(* IEC 61131-3 sources: STAR-PLC-Agent/results/raw/batch_fresh_20261114/PUB003/functional/attempt_0001, 1 file *)

(* ---- test_program.st ---- *)
PROGRAM PLC_PRG
VAR
 BenchStep : UDINT := 0;
 BenchCalls : UDINT := 0;
 BenchDone : BOOL := FALSE;
 BenchUut0 : FB_Task;
 BenchUut1 : FB_Task;
 BenchUut2 : FB_Task;
 BenchUut3 : FB_Task;
 BenchUut4 : FB_Task;
 BenchUut5 : FB_Task;
 BenchUut6 : FB_Task;
 BenchUut7 : FB_Task;
 TraceIn_Value : ARRAY[0..48] OF REAL;
 TraceIn_hiLevel : ARRAY[0..48] OF REAL;
 TraceIn_loLevel : ARRAY[0..48] OF REAL;
 TraceIn_hystWindow : ARRAY[0..48] OF REAL;
 TraceOut_hiAlarm : ARRAY[0..48] OF BOOL;
 TraceOut_loAlarm : ARRAY[0..48] OF BOOL;
 TraceOut_error : ARRAY[0..48] OF BOOL;
 TraceOut_status : ARRAY[0..48] OF WORD;
END_VAR

IF NOT BenchDone THEN
 CASE BenchStep OF
 0:
   BenchUut0.Value := REAL#50.0;
   BenchUut0.hiLevel := REAL#80.0;
   BenchUut0.loLevel := REAL#20.0;
   BenchUut0.hystWindow := REAL#5.0;
   TraceIn_Value[0] := BenchUut0.Value;
   TraceIn_hiLevel[0] := BenchUut0.hiLevel;
   TraceIn_loLevel[0] := BenchUut0.loLevel;
   TraceIn_hystWindow[0] := BenchUut0.hystWindow;
   BenchUut0();
   TraceOut_hiAlarm[0] := BenchUut0.hiAlarm;
   TraceOut_loAlarm[0] := BenchUut0.loAlarm;
   TraceOut_error[0] := BenchUut0.error;
   TraceOut_status[0] := BenchUut0.status;
   BenchCalls := BenchCalls + 1;
 1:
   BenchUut0.Value := REAL#80.0;
   BenchUut0.hiLevel := REAL#80.0;
   BenchUut0.loLevel := REAL#20.0;
   BenchUut0.hystWindow := REAL#5.0;
   TraceIn_Value[1] := BenchUut0.Value;
   TraceIn_hiLevel[1] := BenchUut0.hiLevel;
   TraceIn_loLevel[1] := BenchUut0.loLevel;
   TraceIn_hystWindow[1] := BenchUut0.hystWindow;
   BenchUut0();
   TraceOut_hiAlarm[1] := BenchUut0.hiAlarm;
   TraceOut_loAlarm[1] := BenchUut0.loAlarm;
   TraceOut_error[1] := BenchUut0.error;
   TraceOut_status[1] := BenchUut0.status;
   BenchCalls := BenchCalls + 1;
 2:
   BenchUut0.Value := REAL#81.0;
   BenchUut0.hiLevel := REAL#80.0;
   BenchUut0.loLevel := REAL#20.0;
   BenchUut0.hystWindow := REAL#5.0;
   TraceIn_Value[2] := BenchUut0.Value;
   TraceIn_hiLevel[2] := BenchUut0.hiLevel;
   TraceIn_loLevel[2] := BenchUut0.loLevel;
   TraceIn_hystWindow[2] := BenchUut0.hystWindow;
   BenchUut0();
   TraceOut_hiAlarm[2] := BenchUut0.hiAlarm;
   TraceOut_loAlarm[2] := BenchUut0.loAlarm;
   TraceOut_error[2] := BenchUut0.error;
   TraceOut_status[2] := BenchUut0.status;
   BenchCalls := BenchCalls + 1;
 3:
   BenchUut0.Value := REAL#75.0;
   BenchUut0.hiLevel := REAL#80.0;
   BenchUut0.loLevel := REAL#20.0;
   BenchUut0.hystWindow := REAL#5.0;
   TraceIn_Value[3] := BenchUut0.Value;
   TraceIn_hiLevel[3] := BenchUut0.hiLevel;
   TraceIn_loLevel[3] := BenchUut0.loLevel;
   TraceIn_hystWindow[3] := BenchUut0.hystWindow;
   BenchUut0();
   TraceOut_hiAlarm[3] := BenchUut0.hiAlarm;
   TraceOut_loAlarm[3] := BenchUut0.loAlarm;
   TraceOut_error[3] := BenchUut0.error;
   TraceOut_status[3] := BenchUut0.status;
   BenchCalls := BenchCalls + 1;
 4:
   BenchUut0.Value := REAL#74.0;
   BenchUut0.hiLevel := REAL#80.0;
   BenchUut0.loLevel := REAL#20.0;
   BenchUut0.hystWindow := REAL#5.0;
   TraceIn_Value[4] := BenchUut0.Value;
   TraceIn_hiLevel[4] := BenchUut0.hiLevel;
   TraceIn_loLevel[4] := BenchUut0.loLevel;
   TraceIn_hystWindow[4] := BenchUut0.hystWindow;
   BenchUut0();
   TraceOut_hiAlarm[4] := BenchUut0.hiAlarm;
   TraceOut_loAlarm[4] := BenchUut0.loAlarm;
   TraceOut_error[4] := BenchUut0.error;
   TraceOut_status[4] := BenchUut0.status;
   BenchCalls := BenchCalls + 1;
 5:
   BenchUut0.Value := REAL#20.0;
   BenchUut0.hiLevel := REAL#80.0;
   BenchUut0.loLevel := REAL#20.0;
   BenchUut0.hystWindow := REAL#5.0;
   TraceIn_Value[5] := BenchUut0.Value;
   TraceIn_hiLevel[5] := BenchUut0.hiLevel;
   TraceIn_loLevel[5] := BenchUut0.loLevel;
   TraceIn_hystWindow[5] := BenchUut0.hystWindow;
   BenchUut0();
   TraceOut_hiAlarm[5] := BenchUut0.hiAlarm;
   TraceOut_loAlarm[5] := BenchUut0.loAlarm;
   TraceOut_error[5] := BenchUut0.error;
   TraceOut_status[5] := BenchUut0.status;
   BenchCalls := BenchCalls + 1;
 6:
   BenchUut0.Value := REAL#19.0;
   BenchUut0.hiLevel := REAL#80.0;
   BenchUut0.loLevel := REAL#20.0;
   BenchUut0.hystWindow := REAL#5.0;
   TraceIn_Value[6] := BenchUut0.Value;
   TraceIn_hiLevel[6] := BenchUut0.hiLevel;
   TraceIn_loLevel[6] := BenchUut0.loLevel;
   TraceIn_hystWindow[6] := BenchUut0.hystWindow;
   BenchUut0();
   TraceOut_hiAlarm[6] := BenchUut0.hiAlarm;
   TraceOut_loAlarm[6] := BenchUut0.loAlarm;
   TraceOut_error[6] := BenchUut0.error;
   TraceOut_status[6] := BenchUut0.status;
   BenchCalls := BenchCalls + 1;
 7:
   BenchUut0.Value := REAL#25.0;
   BenchUut0.hiLevel := REAL#80.0;
   BenchUut0.loLevel := REAL#20.0;
   BenchUut0.hystWindow := REAL#5.0;
   TraceIn_Value[7] := BenchUut0.Value;
   TraceIn_hiLevel[7] := BenchUut0.hiLevel;
   TraceIn_loLevel[7] := BenchUut0.loLevel;
   TraceIn_hystWindow[7] := BenchUut0.hystWindow;
   BenchUut0();
   TraceOut_hiAlarm[7] := BenchUut0.hiAlarm;
   TraceOut_loAlarm[7] := BenchUut0.loAlarm;
   TraceOut_error[7] := BenchUut0.error;
   TraceOut_status[7] := BenchUut0.status;
   BenchCalls := BenchCalls + 1;
 8:
   BenchUut0.Value := REAL#26.0;
   BenchUut0.hiLevel := REAL#80.0;
   BenchUut0.loLevel := REAL#20.0;
   BenchUut0.hystWindow := REAL#5.0;
   TraceIn_Value[8] := BenchUut0.Value;
   TraceIn_hiLevel[8] := BenchUut0.hiLevel;
   TraceIn_loLevel[8] := BenchUut0.loLevel;
   TraceIn_hystWindow[8] := BenchUut0.hystWindow;
   BenchUut0();
   TraceOut_hiAlarm[8] := BenchUut0.hiAlarm;
   TraceOut_loAlarm[8] := BenchUut0.loAlarm;
   TraceOut_error[8] := BenchUut0.error;
   TraceOut_status[8] := BenchUut0.status;
   BenchCalls := BenchCalls + 1;
 9:
   BenchUut1.Value := REAL#90.0;
   BenchUut1.hiLevel := REAL#80.0;
   BenchUut1.loLevel := REAL#20.0;
   BenchUut1.hystWindow := REAL#5.0;
   TraceIn_Value[9] := BenchUut1.Value;
   TraceIn_hiLevel[9] := BenchUut1.hiLevel;
   TraceIn_loLevel[9] := BenchUut1.loLevel;
   TraceIn_hystWindow[9] := BenchUut1.hystWindow;
   BenchUut1();
   TraceOut_hiAlarm[9] := BenchUut1.hiAlarm;
   TraceOut_loAlarm[9] := BenchUut1.loAlarm;
   TraceOut_error[9] := BenchUut1.error;
   TraceOut_status[9] := BenchUut1.status;
   BenchCalls := BenchCalls + 1;
 10:
   BenchUut1.Value := REAL#50.0;
   BenchUut1.hiLevel := REAL#80.0;
   BenchUut1.loLevel := REAL#80.0;
   BenchUut1.hystWindow := REAL#80.0;
   TraceIn_Value[10] := BenchUut1.Value;
   TraceIn_hiLevel[10] := BenchUut1.hiLevel;
   TraceIn_loLevel[10] := BenchUut1.loLevel;
   TraceIn_hystWindow[10] := BenchUut1.hystWindow;
   BenchUut1();
   TraceOut_hiAlarm[10] := BenchUut1.hiAlarm;
   TraceOut_loAlarm[10] := BenchUut1.loAlarm;
   TraceOut_error[10] := BenchUut1.error;
   TraceOut_status[10] := BenchUut1.status;
   BenchCalls := BenchCalls + 1;
 11:
   BenchUut1.Value := REAL#50.0;
   BenchUut1.hiLevel := REAL#80.0;
   BenchUut1.loLevel := REAL#20.0;
   BenchUut1.hystWindow := REAL#60.0;
   TraceIn_Value[11] := BenchUut1.Value;
   TraceIn_hiLevel[11] := BenchUut1.hiLevel;
   TraceIn_loLevel[11] := BenchUut1.loLevel;
   TraceIn_hystWindow[11] := BenchUut1.hystWindow;
   BenchUut1();
   TraceOut_hiAlarm[11] := BenchUut1.hiAlarm;
   TraceOut_loAlarm[11] := BenchUut1.loAlarm;
   TraceOut_error[11] := BenchUut1.error;
   TraceOut_status[11] := BenchUut1.status;
   BenchCalls := BenchCalls + 1;
 12:
   BenchUut1.Value := REAL#50.0;
   BenchUut1.hiLevel := REAL#80.0;
   BenchUut1.loLevel := REAL#20.0;
   BenchUut1.hystWindow := REAL#5.0;
   TraceIn_Value[12] := BenchUut1.Value;
   TraceIn_hiLevel[12] := BenchUut1.hiLevel;
   TraceIn_loLevel[12] := BenchUut1.loLevel;
   TraceIn_hystWindow[12] := BenchUut1.hystWindow;
   BenchUut1();
   TraceOut_hiAlarm[12] := BenchUut1.hiAlarm;
   TraceOut_loAlarm[12] := BenchUut1.loAlarm;
   TraceOut_error[12] := BenchUut1.error;
   TraceOut_status[12] := BenchUut1.status;
   BenchCalls := BenchCalls + 1;
 13:
   BenchUut2.Value := REAL#101.0;
   BenchUut2.hiLevel := REAL#100.0;
   BenchUut2.loLevel := REAL#0.0;
   BenchUut2.hystWindow := REAL#90.0;
   TraceIn_Value[13] := BenchUut2.Value;
   TraceIn_hiLevel[13] := BenchUut2.hiLevel;
   TraceIn_loLevel[13] := BenchUut2.loLevel;
   TraceIn_hystWindow[13] := BenchUut2.hystWindow;
   BenchUut2();
   TraceOut_hiAlarm[13] := BenchUut2.hiAlarm;
   TraceOut_loAlarm[13] := BenchUut2.loAlarm;
   TraceOut_error[13] := BenchUut2.error;
   TraceOut_status[13] := BenchUut2.status;
   BenchCalls := BenchCalls + 1;
 14:
   BenchUut2.Value := REAL#50.0;
   BenchUut2.hiLevel := REAL#100.0;
   BenchUut2.loLevel := REAL#0.0;
   BenchUut2.hystWindow := REAL#90.0;
   TraceIn_Value[14] := BenchUut2.Value;
   TraceIn_hiLevel[14] := BenchUut2.hiLevel;
   TraceIn_loLevel[14] := BenchUut2.loLevel;
   TraceIn_hystWindow[14] := BenchUut2.hystWindow;
   BenchUut2();
   TraceOut_hiAlarm[14] := BenchUut2.hiAlarm;
   TraceOut_loAlarm[14] := BenchUut2.loAlarm;
   TraceOut_error[14] := BenchUut2.error;
   TraceOut_status[14] := BenchUut2.status;
   BenchCalls := BenchCalls + 1;
 15:
   BenchUut2.Value := REAL#50.0;
   BenchUut2.hiLevel := REAL#100.0;
   BenchUut2.loLevel := REAL#100.0;
   BenchUut2.hystWindow := REAL#90.0;
   TraceIn_Value[15] := BenchUut2.Value;
   TraceIn_hiLevel[15] := BenchUut2.hiLevel;
   TraceIn_loLevel[15] := BenchUut2.loLevel;
   TraceIn_hystWindow[15] := BenchUut2.hystWindow;
   BenchUut2();
   TraceOut_hiAlarm[15] := BenchUut2.hiAlarm;
   TraceOut_loAlarm[15] := BenchUut2.loAlarm;
   TraceOut_error[15] := BenchUut2.error;
   TraceOut_status[15] := BenchUut2.status;
   BenchCalls := BenchCalls + 1;
 16:
   BenchUut2.Value := REAL#10.0;
   BenchUut2.hiLevel := REAL#100.0;
   BenchUut2.loLevel := REAL#0.0;
   BenchUut2.hystWindow := REAL#90.0;
   TraceIn_Value[16] := BenchUut2.Value;
   TraceIn_hiLevel[16] := BenchUut2.hiLevel;
   TraceIn_loLevel[16] := BenchUut2.loLevel;
   TraceIn_hystWindow[16] := BenchUut2.hystWindow;
   BenchUut2();
   TraceOut_hiAlarm[16] := BenchUut2.hiAlarm;
   TraceOut_loAlarm[16] := BenchUut2.loAlarm;
   TraceOut_error[16] := BenchUut2.error;
   TraceOut_status[16] := BenchUut2.status;
   BenchCalls := BenchCalls + 1;
 17:
   BenchUut2.Value := REAL#9.0;
   BenchUut2.hiLevel := REAL#100.0;
   BenchUut2.loLevel := REAL#0.0;
   BenchUut2.hystWindow := REAL#90.0;
   TraceIn_Value[17] := BenchUut2.Value;
   TraceIn_hiLevel[17] := BenchUut2.hiLevel;
   TraceIn_loLevel[17] := BenchUut2.loLevel;
   TraceIn_hystWindow[17] := BenchUut2.hystWindow;
   BenchUut2();
   TraceOut_hiAlarm[17] := BenchUut2.hiAlarm;
   TraceOut_loAlarm[17] := BenchUut2.loAlarm;
   TraceOut_error[17] := BenchUut2.error;
   TraceOut_status[17] := BenchUut2.status;
   BenchCalls := BenchCalls + 1;
 18:
   BenchUut2.Value := REAL#-1.0;
   BenchUut2.hiLevel := REAL#100.0;
   BenchUut2.loLevel := REAL#0.0;
   BenchUut2.hystWindow := REAL#90.0;
   TraceIn_Value[18] := BenchUut2.Value;
   TraceIn_hiLevel[18] := BenchUut2.hiLevel;
   TraceIn_loLevel[18] := BenchUut2.loLevel;
   TraceIn_hystWindow[18] := BenchUut2.hystWindow;
   BenchUut2();
   TraceOut_hiAlarm[18] := BenchUut2.hiAlarm;
   TraceOut_loAlarm[18] := BenchUut2.loAlarm;
   TraceOut_error[18] := BenchUut2.error;
   TraceOut_status[18] := BenchUut2.status;
   BenchCalls := BenchCalls + 1;
 19:
   BenchUut3.Value := REAL#5.0;
   BenchUut3.hiLevel := REAL#50.0;
   BenchUut3.loLevel := REAL#10.0;
   BenchUut3.hystWindow := REAL#5.0;
   TraceIn_Value[19] := BenchUut3.Value;
   TraceIn_hiLevel[19] := BenchUut3.hiLevel;
   TraceIn_loLevel[19] := BenchUut3.loLevel;
   TraceIn_hystWindow[19] := BenchUut3.hystWindow;
   BenchUut3();
   TraceOut_hiAlarm[19] := BenchUut3.hiAlarm;
   TraceOut_loAlarm[19] := BenchUut3.loAlarm;
   TraceOut_error[19] := BenchUut3.error;
   TraceOut_status[19] := BenchUut3.status;
   BenchCalls := BenchCalls + 1;
 20:
   BenchUut3.Value := REAL#25.0;
   BenchUut3.hiLevel := REAL#50.0;
   BenchUut3.loLevel := REAL#60.0;
   BenchUut3.hystWindow := REAL#5.0;
   TraceIn_Value[20] := BenchUut3.Value;
   TraceIn_hiLevel[20] := BenchUut3.hiLevel;
   TraceIn_loLevel[20] := BenchUut3.loLevel;
   TraceIn_hystWindow[20] := BenchUut3.hystWindow;
   BenchUut3();
   TraceOut_hiAlarm[20] := BenchUut3.hiAlarm;
   TraceOut_loAlarm[20] := BenchUut3.loAlarm;
   TraceOut_error[20] := BenchUut3.error;
   TraceOut_status[20] := BenchUut3.status;
   BenchCalls := BenchCalls + 1;
 21:
   BenchUut3.Value := REAL#25.0;
   BenchUut3.hiLevel := REAL#50.0;
   BenchUut3.loLevel := REAL#10.0;
   BenchUut3.hystWindow := REAL#40.0;
   TraceIn_Value[21] := BenchUut3.Value;
   TraceIn_hiLevel[21] := BenchUut3.hiLevel;
   TraceIn_loLevel[21] := BenchUut3.loLevel;
   TraceIn_hystWindow[21] := BenchUut3.hystWindow;
   BenchUut3();
   TraceOut_hiAlarm[21] := BenchUut3.hiAlarm;
   TraceOut_loAlarm[21] := BenchUut3.loAlarm;
   TraceOut_error[21] := BenchUut3.error;
   TraceOut_status[21] := BenchUut3.status;
   BenchCalls := BenchCalls + 1;
 22:
   BenchUut3.Value := REAL#16.0;
   BenchUut3.hiLevel := REAL#50.0;
   BenchUut3.loLevel := REAL#10.0;
   BenchUut3.hystWindow := REAL#5.0;
   TraceIn_Value[22] := BenchUut3.Value;
   TraceIn_hiLevel[22] := BenchUut3.hiLevel;
   TraceIn_loLevel[22] := BenchUut3.loLevel;
   TraceIn_hystWindow[22] := BenchUut3.hystWindow;
   BenchUut3();
   TraceOut_hiAlarm[22] := BenchUut3.hiAlarm;
   TraceOut_loAlarm[22] := BenchUut3.loAlarm;
   TraceOut_error[22] := BenchUut3.error;
   TraceOut_status[22] := BenchUut3.status;
   BenchCalls := BenchCalls + 1;
 23:
   BenchUut3.Value := REAL#10.125;
   BenchUut3.hiLevel := REAL#20.375;
   BenchUut3.loLevel := REAL#10.125;
   BenchUut3.hystWindow := REAL#0.0;
   TraceIn_Value[23] := BenchUut3.Value;
   TraceIn_hiLevel[23] := BenchUut3.hiLevel;
   TraceIn_loLevel[23] := BenchUut3.loLevel;
   TraceIn_hystWindow[23] := BenchUut3.hystWindow;
   BenchUut3();
   TraceOut_hiAlarm[23] := BenchUut3.hiAlarm;
   TraceOut_loAlarm[23] := BenchUut3.loAlarm;
   TraceOut_error[23] := BenchUut3.error;
   TraceOut_status[23] := BenchUut3.status;
   BenchCalls := BenchCalls + 1;
 24:
   BenchUut3.Value := REAL#20.3751;
   BenchUut3.hiLevel := REAL#20.375;
   BenchUut3.loLevel := REAL#10.125;
   BenchUut3.hystWindow := REAL#0.0;
   TraceIn_Value[24] := BenchUut3.Value;
   TraceIn_hiLevel[24] := BenchUut3.hiLevel;
   TraceIn_loLevel[24] := BenchUut3.loLevel;
   TraceIn_hystWindow[24] := BenchUut3.hystWindow;
   BenchUut3();
   TraceOut_hiAlarm[24] := BenchUut3.hiAlarm;
   TraceOut_loAlarm[24] := BenchUut3.loAlarm;
   TraceOut_error[24] := BenchUut3.error;
   TraceOut_status[24] := BenchUut3.status;
   BenchCalls := BenchCalls + 1;
 25:
   BenchUut3.Value := REAL#20.25;
   BenchUut3.hiLevel := REAL#20.375;
   BenchUut3.loLevel := REAL#10.125;
   BenchUut3.hystWindow := REAL#0.0;
   TraceIn_Value[25] := BenchUut3.Value;
   TraceIn_hiLevel[25] := BenchUut3.hiLevel;
   TraceIn_loLevel[25] := BenchUut3.loLevel;
   TraceIn_hystWindow[25] := BenchUut3.hystWindow;
   BenchUut3();
   TraceOut_hiAlarm[25] := BenchUut3.hiAlarm;
   TraceOut_loAlarm[25] := BenchUut3.loAlarm;
   TraceOut_error[25] := BenchUut3.error;
   TraceOut_status[25] := BenchUut3.status;
   BenchCalls := BenchCalls + 1;
 26:
   BenchUut4.Value := REAL#19.0;
   BenchUut4.hiLevel := REAL#80.0;
   BenchUut4.loLevel := REAL#20.0;
   BenchUut4.hystWindow := REAL#5.0;
   TraceIn_Value[26] := BenchUut4.Value;
   TraceIn_hiLevel[26] := BenchUut4.hiLevel;
   TraceIn_loLevel[26] := BenchUut4.loLevel;
   TraceIn_hystWindow[26] := BenchUut4.hystWindow;
   BenchUut4();
   TraceOut_hiAlarm[26] := BenchUut4.hiAlarm;
   TraceOut_loAlarm[26] := BenchUut4.loAlarm;
   TraceOut_error[26] := BenchUut4.error;
   TraceOut_status[26] := BenchUut4.status;
   BenchCalls := BenchCalls + 1;
 27:
   BenchUut4.Value := REAL#50.0;
   BenchUut4.hiLevel := REAL#80.0;
   BenchUut4.loLevel := REAL#80.0;
   BenchUut4.hystWindow := REAL#80.0;
   TraceIn_Value[27] := BenchUut4.Value;
   TraceIn_hiLevel[27] := BenchUut4.hiLevel;
   TraceIn_loLevel[27] := BenchUut4.loLevel;
   TraceIn_hystWindow[27] := BenchUut4.hystWindow;
   BenchUut4();
   TraceOut_hiAlarm[27] := BenchUut4.hiAlarm;
   TraceOut_loAlarm[27] := BenchUut4.loAlarm;
   TraceOut_error[27] := BenchUut4.error;
   TraceOut_status[27] := BenchUut4.status;
   BenchCalls := BenchCalls + 1;
 28:
   BenchUut5.Value := REAL#1.1;
   BenchUut5.hiLevel := REAL#1.0;
   BenchUut5.loLevel := REAL#0.0;
   BenchUut5.hystWindow := REAL#0.10000000149011612;
   TraceIn_Value[28] := BenchUut5.Value;
   TraceIn_hiLevel[28] := BenchUut5.hiLevel;
   TraceIn_loLevel[28] := BenchUut5.loLevel;
   TraceIn_hystWindow[28] := BenchUut5.hystWindow;
   BenchUut5();
   TraceOut_hiAlarm[28] := BenchUut5.hiAlarm;
   TraceOut_loAlarm[28] := BenchUut5.loAlarm;
   TraceOut_error[28] := BenchUut5.error;
   TraceOut_status[28] := BenchUut5.status;
   BenchCalls := BenchCalls + 1;
 29:
   BenchUut5.Value := REAL#1.0;
   BenchUut5.hiLevel := REAL#1.0;
   BenchUut5.loLevel := REAL#0.0;
   BenchUut5.hystWindow := REAL#0.10000000149011612;
   TraceIn_Value[29] := BenchUut5.Value;
   TraceIn_hiLevel[29] := BenchUut5.hiLevel;
   TraceIn_loLevel[29] := BenchUut5.loLevel;
   TraceIn_hystWindow[29] := BenchUut5.hystWindow;
   BenchUut5();
   TraceOut_hiAlarm[29] := BenchUut5.hiAlarm;
   TraceOut_loAlarm[29] := BenchUut5.loAlarm;
   TraceOut_error[29] := BenchUut5.error;
   TraceOut_status[29] := BenchUut5.status;
   BenchCalls := BenchCalls + 1;
 30:
   BenchUut5.Value := REAL#0.8999999761581421;
   BenchUut5.hiLevel := REAL#1.0;
   BenchUut5.loLevel := REAL#0.0;
   BenchUut5.hystWindow := REAL#0.10000000149011612;
   TraceIn_Value[30] := BenchUut5.Value;
   TraceIn_hiLevel[30] := BenchUut5.hiLevel;
   TraceIn_loLevel[30] := BenchUut5.loLevel;
   TraceIn_hystWindow[30] := BenchUut5.hystWindow;
   BenchUut5();
   TraceOut_hiAlarm[30] := BenchUut5.hiAlarm;
   TraceOut_loAlarm[30] := BenchUut5.loAlarm;
   TraceOut_error[30] := BenchUut5.error;
   TraceOut_status[30] := BenchUut5.status;
   BenchCalls := BenchCalls + 1;
 31:
   BenchUut5.Value := REAL#0.8999989628791809;
   BenchUut5.hiLevel := REAL#1.0;
   BenchUut5.loLevel := REAL#0.0;
   BenchUut5.hystWindow := REAL#0.10000000149011612;
   TraceIn_Value[31] := BenchUut5.Value;
   TraceIn_hiLevel[31] := BenchUut5.hiLevel;
   TraceIn_loLevel[31] := BenchUut5.loLevel;
   TraceIn_hystWindow[31] := BenchUut5.hystWindow;
   BenchUut5();
   TraceOut_hiAlarm[31] := BenchUut5.hiAlarm;
   TraceOut_loAlarm[31] := BenchUut5.loAlarm;
   TraceOut_error[31] := BenchUut5.error;
   TraceOut_status[31] := BenchUut5.status;
   BenchCalls := BenchCalls + 1;
 32:
   BenchUut5.Value := REAL#-0.1;
   BenchUut5.hiLevel := REAL#1.0;
   BenchUut5.loLevel := REAL#0.0;
   BenchUut5.hystWindow := REAL#0.10000000149011612;
   TraceIn_Value[32] := BenchUut5.Value;
   TraceIn_hiLevel[32] := BenchUut5.hiLevel;
   TraceIn_loLevel[32] := BenchUut5.loLevel;
   TraceIn_hystWindow[32] := BenchUut5.hystWindow;
   BenchUut5();
   TraceOut_hiAlarm[32] := BenchUut5.hiAlarm;
   TraceOut_loAlarm[32] := BenchUut5.loAlarm;
   TraceOut_error[32] := BenchUut5.error;
   TraceOut_status[32] := BenchUut5.status;
   BenchCalls := BenchCalls + 1;
 33:
   BenchUut5.Value := REAL#0.0;
   BenchUut5.hiLevel := REAL#1.0;
   BenchUut5.loLevel := REAL#0.0;
   BenchUut5.hystWindow := REAL#0.10000000149011612;
   TraceIn_Value[33] := BenchUut5.Value;
   TraceIn_hiLevel[33] := BenchUut5.hiLevel;
   TraceIn_loLevel[33] := BenchUut5.loLevel;
   TraceIn_hystWindow[33] := BenchUut5.hystWindow;
   BenchUut5();
   TraceOut_hiAlarm[33] := BenchUut5.hiAlarm;
   TraceOut_loAlarm[33] := BenchUut5.loAlarm;
   TraceOut_error[33] := BenchUut5.error;
   TraceOut_status[33] := BenchUut5.status;
   BenchCalls := BenchCalls + 1;
 34:
   BenchUut5.Value := REAL#0.10000000149011612;
   BenchUut5.hiLevel := REAL#1.0;
   BenchUut5.loLevel := REAL#0.0;
   BenchUut5.hystWindow := REAL#0.10000000149011612;
   TraceIn_Value[34] := BenchUut5.Value;
   TraceIn_hiLevel[34] := BenchUut5.hiLevel;
   TraceIn_loLevel[34] := BenchUut5.loLevel;
   TraceIn_hystWindow[34] := BenchUut5.hystWindow;
   BenchUut5();
   TraceOut_hiAlarm[34] := BenchUut5.hiAlarm;
   TraceOut_loAlarm[34] := BenchUut5.loAlarm;
   TraceOut_error[34] := BenchUut5.error;
   TraceOut_status[34] := BenchUut5.status;
   BenchCalls := BenchCalls + 1;
 35:
   BenchUut5.Value := REAL#0.10000099986791611;
   BenchUut5.hiLevel := REAL#1.0;
   BenchUut5.loLevel := REAL#0.0;
   BenchUut5.hystWindow := REAL#0.10000000149011612;
   TraceIn_Value[35] := BenchUut5.Value;
   TraceIn_hiLevel[35] := BenchUut5.hiLevel;
   TraceIn_loLevel[35] := BenchUut5.loLevel;
   TraceIn_hystWindow[35] := BenchUut5.hystWindow;
   BenchUut5();
   TraceOut_hiAlarm[35] := BenchUut5.hiAlarm;
   TraceOut_loAlarm[35] := BenchUut5.loAlarm;
   TraceOut_error[35] := BenchUut5.error;
   TraceOut_status[35] := BenchUut5.status;
   BenchCalls := BenchCalls + 1;
 36:
   BenchUut6.Value := REAL#-9.0;
   BenchUut6.hiLevel := REAL#-10.0;
   BenchUut6.loLevel := REAL#-50.0;
   BenchUut6.hystWindow := REAL#5.0;
   TraceIn_Value[36] := BenchUut6.Value;
   TraceIn_hiLevel[36] := BenchUut6.hiLevel;
   TraceIn_loLevel[36] := BenchUut6.loLevel;
   TraceIn_hystWindow[36] := BenchUut6.hystWindow;
   BenchUut6();
   TraceOut_hiAlarm[36] := BenchUut6.hiAlarm;
   TraceOut_loAlarm[36] := BenchUut6.loAlarm;
   TraceOut_error[36] := BenchUut6.error;
   TraceOut_status[36] := BenchUut6.status;
   BenchCalls := BenchCalls + 1;
 37:
   BenchUut6.Value := REAL#-15.0;
   BenchUut6.hiLevel := REAL#-10.0;
   BenchUut6.loLevel := REAL#-50.0;
   BenchUut6.hystWindow := REAL#5.0;
   TraceIn_Value[37] := BenchUut6.Value;
   TraceIn_hiLevel[37] := BenchUut6.hiLevel;
   TraceIn_loLevel[37] := BenchUut6.loLevel;
   TraceIn_hystWindow[37] := BenchUut6.hystWindow;
   BenchUut6();
   TraceOut_hiAlarm[37] := BenchUut6.hiAlarm;
   TraceOut_loAlarm[37] := BenchUut6.loAlarm;
   TraceOut_error[37] := BenchUut6.error;
   TraceOut_status[37] := BenchUut6.status;
   BenchCalls := BenchCalls + 1;
 38:
   BenchUut6.Value := REAL#-15.1;
   BenchUut6.hiLevel := REAL#-10.0;
   BenchUut6.loLevel := REAL#-50.0;
   BenchUut6.hystWindow := REAL#5.0;
   TraceIn_Value[38] := BenchUut6.Value;
   TraceIn_hiLevel[38] := BenchUut6.hiLevel;
   TraceIn_loLevel[38] := BenchUut6.loLevel;
   TraceIn_hystWindow[38] := BenchUut6.hystWindow;
   BenchUut6();
   TraceOut_hiAlarm[38] := BenchUut6.hiAlarm;
   TraceOut_loAlarm[38] := BenchUut6.loAlarm;
   TraceOut_error[38] := BenchUut6.error;
   TraceOut_status[38] := BenchUut6.status;
   BenchCalls := BenchCalls + 1;
 39:
   BenchUut6.Value := REAL#-51.0;
   BenchUut6.hiLevel := REAL#-10.0;
   BenchUut6.loLevel := REAL#-50.0;
   BenchUut6.hystWindow := REAL#5.0;
   TraceIn_Value[39] := BenchUut6.Value;
   TraceIn_hiLevel[39] := BenchUut6.hiLevel;
   TraceIn_loLevel[39] := BenchUut6.loLevel;
   TraceIn_hystWindow[39] := BenchUut6.hystWindow;
   BenchUut6();
   TraceOut_hiAlarm[39] := BenchUut6.hiAlarm;
   TraceOut_loAlarm[39] := BenchUut6.loAlarm;
   TraceOut_error[39] := BenchUut6.error;
   TraceOut_status[39] := BenchUut6.status;
   BenchCalls := BenchCalls + 1;
 40:
   BenchUut6.Value := REAL#-45.0;
   BenchUut6.hiLevel := REAL#-10.0;
   BenchUut6.loLevel := REAL#-50.0;
   BenchUut6.hystWindow := REAL#5.0;
   TraceIn_Value[40] := BenchUut6.Value;
   TraceIn_hiLevel[40] := BenchUut6.hiLevel;
   TraceIn_loLevel[40] := BenchUut6.loLevel;
   TraceIn_hystWindow[40] := BenchUut6.hystWindow;
   BenchUut6();
   TraceOut_hiAlarm[40] := BenchUut6.hiAlarm;
   TraceOut_loAlarm[40] := BenchUut6.loAlarm;
   TraceOut_error[40] := BenchUut6.error;
   TraceOut_status[40] := BenchUut6.status;
   BenchCalls := BenchCalls + 1;
 41:
   BenchUut6.Value := REAL#-44.9;
   BenchUut6.hiLevel := REAL#-10.0;
   BenchUut6.loLevel := REAL#-50.0;
   BenchUut6.hystWindow := REAL#5.0;
   TraceIn_Value[41] := BenchUut6.Value;
   TraceIn_hiLevel[41] := BenchUut6.hiLevel;
   TraceIn_loLevel[41] := BenchUut6.loLevel;
   TraceIn_hystWindow[41] := BenchUut6.hystWindow;
   BenchUut6();
   TraceOut_hiAlarm[41] := BenchUut6.hiAlarm;
   TraceOut_loAlarm[41] := BenchUut6.loAlarm;
   TraceOut_error[41] := BenchUut6.error;
   TraceOut_status[41] := BenchUut6.status;
   BenchCalls := BenchCalls + 1;
 42:
   BenchUut6.Value := REAL#0.0;
   BenchUut6.hiLevel := REAL#-10.0;
   BenchUut6.loLevel := REAL#-50.0;
   BenchUut6.hystWindow := REAL#5.0;
   TraceIn_Value[42] := BenchUut6.Value;
   TraceIn_hiLevel[42] := BenchUut6.hiLevel;
   TraceIn_loLevel[42] := BenchUut6.loLevel;
   TraceIn_hystWindow[42] := BenchUut6.hystWindow;
   BenchUut6();
   TraceOut_hiAlarm[42] := BenchUut6.hiAlarm;
   TraceOut_loAlarm[42] := BenchUut6.loAlarm;
   TraceOut_error[42] := BenchUut6.error;
   TraceOut_status[42] := BenchUut6.status;
   BenchCalls := BenchCalls + 1;
 43:
   BenchUut6.Value := REAL#-60.0;
   BenchUut6.hiLevel := REAL#-10.0;
   BenchUut6.loLevel := REAL#-50.0;
   BenchUut6.hystWindow := REAL#5.0;
   TraceIn_Value[43] := BenchUut6.Value;
   TraceIn_hiLevel[43] := BenchUut6.hiLevel;
   TraceIn_loLevel[43] := BenchUut6.loLevel;
   TraceIn_hystWindow[43] := BenchUut6.hystWindow;
   BenchUut6();
   TraceOut_hiAlarm[43] := BenchUut6.hiAlarm;
   TraceOut_loAlarm[43] := BenchUut6.loAlarm;
   TraceOut_error[43] := BenchUut6.error;
   TraceOut_status[43] := BenchUut6.status;
   BenchCalls := BenchCalls + 1;
 44:
   BenchUut7.Value := REAL#85.0;
   BenchUut7.hiLevel := REAL#80.0;
   BenchUut7.loLevel := REAL#20.0;
   BenchUut7.hystWindow := REAL#5.0;
   TraceIn_Value[44] := BenchUut7.Value;
   TraceIn_hiLevel[44] := BenchUut7.hiLevel;
   TraceIn_loLevel[44] := BenchUut7.loLevel;
   TraceIn_hystWindow[44] := BenchUut7.hystWindow;
   BenchUut7();
   TraceOut_hiAlarm[44] := BenchUut7.hiAlarm;
   TraceOut_loAlarm[44] := BenchUut7.loAlarm;
   TraceOut_error[44] := BenchUut7.error;
   TraceOut_status[44] := BenchUut7.status;
   BenchCalls := BenchCalls + 1;
 45:
   BenchUut7.Value := REAL#10.0;
   BenchUut7.hiLevel := REAL#80.0;
   BenchUut7.loLevel := REAL#20.0;
   BenchUut7.hystWindow := REAL#60.0;
   TraceIn_Value[45] := BenchUut7.Value;
   TraceIn_hiLevel[45] := BenchUut7.hiLevel;
   TraceIn_loLevel[45] := BenchUut7.loLevel;
   TraceIn_hystWindow[45] := BenchUut7.hystWindow;
   BenchUut7();
   TraceOut_hiAlarm[45] := BenchUut7.hiAlarm;
   TraceOut_loAlarm[45] := BenchUut7.loAlarm;
   TraceOut_error[45] := BenchUut7.error;
   TraceOut_status[45] := BenchUut7.status;
   BenchCalls := BenchCalls + 1;
 46:
   BenchUut7.Value := REAL#10.0;
   BenchUut7.hiLevel := REAL#50.0;
   BenchUut7.loLevel := REAL#60.0;
   BenchUut7.hystWindow := REAL#5.0;
   TraceIn_Value[46] := BenchUut7.Value;
   TraceIn_hiLevel[46] := BenchUut7.hiLevel;
   TraceIn_loLevel[46] := BenchUut7.loLevel;
   TraceIn_hystWindow[46] := BenchUut7.hystWindow;
   BenchUut7();
   TraceOut_hiAlarm[46] := BenchUut7.hiAlarm;
   TraceOut_loAlarm[46] := BenchUut7.loAlarm;
   TraceOut_error[46] := BenchUut7.error;
   TraceOut_status[46] := BenchUut7.status;
   BenchCalls := BenchCalls + 1;
 47:
   BenchUut7.Value := REAL#75.0;
   BenchUut7.hiLevel := REAL#80.0;
   BenchUut7.loLevel := REAL#20.0;
   BenchUut7.hystWindow := REAL#5.0;
   TraceIn_Value[47] := BenchUut7.Value;
   TraceIn_hiLevel[47] := BenchUut7.hiLevel;
   TraceIn_loLevel[47] := BenchUut7.loLevel;
   TraceIn_hystWindow[47] := BenchUut7.hystWindow;
   BenchUut7();
   TraceOut_hiAlarm[47] := BenchUut7.hiAlarm;
   TraceOut_loAlarm[47] := BenchUut7.loAlarm;
   TraceOut_error[47] := BenchUut7.error;
   TraceOut_status[47] := BenchUut7.status;
   BenchCalls := BenchCalls + 1;
 48:
   BenchUut7.Value := REAL#74.0;
   BenchUut7.hiLevel := REAL#80.0;
   BenchUut7.loLevel := REAL#20.0;
   BenchUut7.hystWindow := REAL#5.0;
   TraceIn_Value[48] := BenchUut7.Value;
   TraceIn_hiLevel[48] := BenchUut7.hiLevel;
   TraceIn_loLevel[48] := BenchUut7.loLevel;
   TraceIn_hystWindow[48] := BenchUut7.hystWindow;
   BenchUut7();
   TraceOut_hiAlarm[48] := BenchUut7.hiAlarm;
   TraceOut_loAlarm[48] := BenchUut7.loAlarm;
   TraceOut_error[48] := BenchUut7.error;
   TraceOut_status[48] := BenchUut7.status;
   BenchCalls := BenchCalls + 1;
 END_CASE;
 BenchStep := BenchStep + 1;
 IF BenchStep >= 49 THEN BenchDone := TRUE; END_IF;
END_IF;
END_PROGRAM
